// TIA Portal V19 export
VAR_GLOBAL   // PLC tag table "R1_OUT"
   "ByteOUT :0 R1" AT %QB78 : Byte;   // System Bits 1
   "ByteOUT :1 R1" AT %QB79 : Byte;   // System Bits 2
   "ByteOUT :2 R1" AT %QB80 : Byte;   // Signals
   "ByteOUT :3 R1" AT %QB81 : Byte;   // Signals
   "ByteOUT :4 R1" AT %QB82 : Byte;   // CMD
   "ByteOUT :5 R1" AT %QB83 : Byte;   // CMD
   "ByteOUT :6 R1" AT %QB84 : Byte;   // X
   "ByteOUT :7 R1" AT %QB85 : Byte;   // X
   "ByteOUT :8 R1" AT %QB86 : Byte;   // Y
   "ByteOUT :9 R1" AT %QB87 : Byte;   // Y
   "ByteOUT :10 R1" AT %QB88 : Byte;   // Z
   "ByteOUT :11 R1" AT %QB89 : Byte;   // Z
   "ByteOUT :12 R1" AT %QB90 : Byte;
   "ByteOUT :13 R1" AT %QB91 : Byte;
   "ByteOUT :14 R1" AT %QB92 : Byte;
   "ByteOUT :15 R1" AT %QB93 : Byte;
   "ByteOUT :16 R1" AT %QB94 : Byte;
   "ByteOUT :17 R1" AT %QB95 : Byte;
   "ByteOUT :18 R1" AT %QB96 : Byte;
   "ByteOUT :19 R1" AT %QB97 : Byte;
   "ByteOUT :20 R1" AT %QB98 : Byte;
   "ByteOUT :21 R1" AT %QB99 : Byte;
   "ByteOUT :22 R1" AT %QB100 : Byte;
   "ByteOUT :23 R1" AT %QB101 : Byte;
   "ByteOUT :24 R1" AT %QB102 : Byte;
   "ByteOUT :25 R1" AT %QB103 : Byte;
   "ByteOUT :26 R1" AT %QB104 : Byte;
   "ByteOUT :27 R1" AT %QB105 : Byte;
   "ByteOUT :28 R1" AT %QB106 : Byte;
   "ByteOUT :29 R1" AT %QB107 : Byte;
   "ByteOUT :30 R1" AT %QB108 : Byte;
   "ByteOUT :31 R1" AT %QB109 : Byte;
   "ByteOUT :32 R1" AT %QB110 : Byte;
   "ByteOUT :33 R1" AT %QB111 : Byte;
   "ByteOUT :34 R1" AT %QB112 : Byte;
   "ByteOUT :35 R1" AT %QB113 : Byte;
   "ByteOUT :36 R1" AT %QB114 : Byte;
   "ByteOUT :37 R1" AT %QB115 : Byte;
   "ByteOUT :38 R1" AT %QB116 : Byte;
   "ByteOUT :39 R1" AT %QB117 : Byte;
   "ByteOUT :40 R1" AT %QB118 : Byte;
   "ByteOUT :41 R1" AT %QB119 : Byte;
   "ByteOUT :42 R1" AT %QB120 : Byte;
   "ByteOUT :43 R1" AT %QB121 : Byte;
   "ByteOUT :44 R1" AT %QB122 : Byte;
   "ByteOUT :45 R1" AT %QB123 : Byte;
   "ByteOUT :46 R1" AT %QB124 : Byte;
   "ByteOUT :47 R1" AT %QB125 : Byte;
   "ByteOUT :48 R1" AT %QB126 : Byte;
   "ByteOUT :49 R1" AT %QB127 : Byte;
   "ByteOUT :50 R1" AT %QB128 : Byte;
   "ByteOUT :51 R1" AT %QB129 : Byte;
   "ByteOUT :52 R1" AT %QB130 : Byte;
   "ByteOUT :53 R1" AT %QB131 : Byte;
   "ByteOUT :54 R1" AT %QB132 : Byte;
   "ByteOUT :55 R1" AT %QB133 : Byte;
   "ByteOUT :56 R1" AT %QB134 : Byte;
   "ByteOUT :57 R1" AT %QB135 : Byte;
   "ByteOUT :58 R1" AT %QB136 : Byte;
   "ByteOUT :59 R1" AT %QB137 : Byte;
   "ByteOUT :60 R1" AT %QB138 : Byte;
   "ByteOUT :61 R1" AT %QB139 : Byte;
   "ByteOUT :62 R1" AT %QB140 : Byte;
   "ByteOUT :63 R1" AT %QB141 : Byte;
END_VAR
